(* IEC 61131-3 sources: codesys-to-s7/tests/corpus/C2S7-TYPE-DATE/neg, 1 file *)

(* ---- input.st ---- *)
FUNCTION_BLOCK FB_Case
VAR
    dtNow : DT;
END_VAR
dtNow := DT#2024-01-01-00:00:00;
END_FUNCTION_BLOCK
